Fanuc KAREL source: compact_preamble.KL

PROGRAM KB00041
%NOLOCKGROUP
VAR
P1 : STRING[80];P2:REAL
BEGIN
P1='A'
P2=1.0
CNV_STR_REAL(P1,P2)
END KB00041
